(* Facility Management Airconditioning Control *)

PROGRAM main
  VAR
    StartButton AT %IX0.0 : BOOL;
    StopButton AT %IX0.1 : BOOL;
    Process AT %MX0.0 : BOOL;
    RoomHot AT %MX0.1 : BOOL;
    AirCon AT %QX0.1 : BOOL;
    MeasuredTemp AT %IW0 : INT;
    ThresholdTemp : INT := 21;
  END_VAR

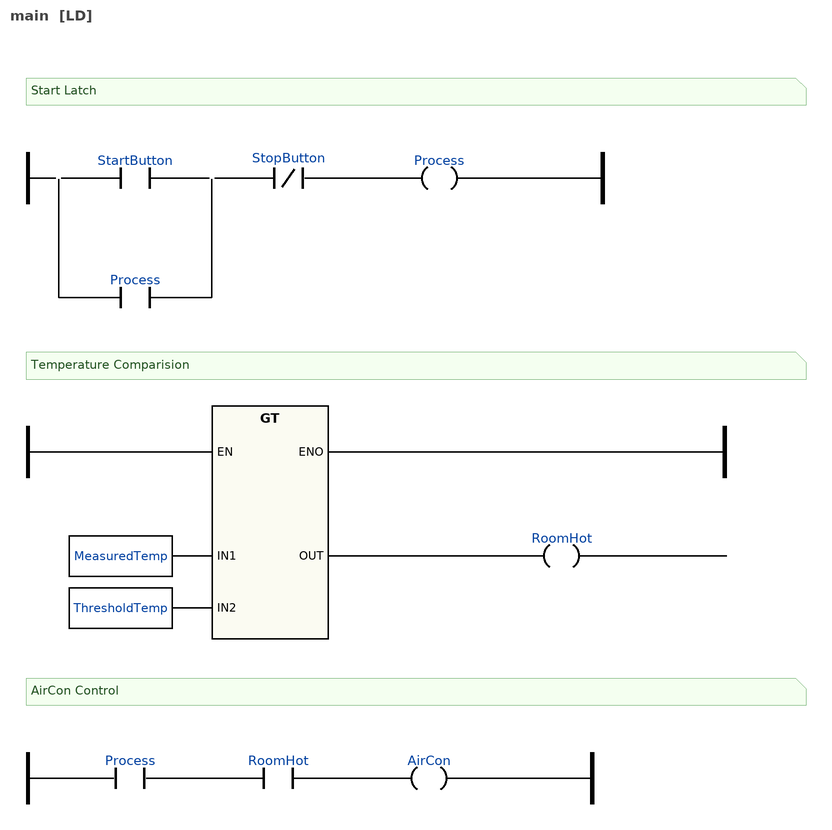
(* LD diagram, written out as Structured Text *)
(* Start Latch *)
Process := (StartButton OR Process) AND NOT StopButton;
(* Temperature Comparision *)
RoomHot := MeasuredTemp > ThresholdTemp;
(* AirCon Control *)
AirCon := Process AND RoomHot;
END_PROGRAM
